ABB RAPID module: LongProg_1.mod

%%%
  VERSION:1
  LANGUAGE:ENGLISH
%%%
MODULE MOD_Tmp2

	PROC Prg_Tmp2()

		MoveAbsJ [[30.000000,25.000000,80.000000,-45.000000,0.000000,0.000000],[9E+09,9E+09,9E+09,9E+09,9E+09,9E+09]],v500,z1,ToolS \WObj:=FrameS;
		MoveAbsJ [[10.000000,-20.000000,50.000000,30.000000,0.000000,0.000000],[9E+09,9E+09,9E+09,9E+09,9E+09,9E+09]],v500,z1,ToolS \WObj:=FrameS;
		MoveAbsJ [[30.000000,25.000000,80.000000,-45.000000,0.000000,0.000000],[9E+09,9E+09,9E+09,9E+09,9E+09,9E+09]],v500,z1,ToolS \WObj:=FrameS;
		MoveAbsJ [[10.000000,-20.000000,50.000000,30.000000,0.000000,0.000000],[9E+09,9E+09,9E+09,9E+09,9E+09,9E+09]],v500,z1,ToolS \WObj:=FrameS;
		MoveAbsJ [[30.000000,25.000000,80.000000,-45.000000,0.000000,0.000000],[9E+09,9E+09,9E+09,9E+09,9E+09,9E+09]],v500,z1,ToolS \WObj:=FrameS;

	ENDPROC

ENDMODULE
